// TIA Portal V20 export
TYPE "Afag_Variablen_Steuerung_Dreh"
   STRUCT
      BA_Manuell : Bool;
      Manuell_Geschwindigkeit_in_P : Int := 10;
      Richten_Reset_FRG : Bool;
      drive_enable : Bool;
      start_homing : Bool;
      jog_pos : Bool;
      jog_neg : Bool;
      fault_reset : Bool;
      Tipp_pos : Bool;
      Tipp_neg : Bool;
      Start_pos_man : Bool;
      Verfahrweg_Grad : Real;
      soll_wert_man_Grad : Real;
      Softw_ES_min_Grad : Real;
      Softw_ES_max_Grad : Real;
      Max_Speed_Grad_s : Real;
      Max_Beschleunigung_Grad_s : Real;
      drive_enable_ok : Bool;
      home_valid : Bool;
      pos_ok : Bool;
      velo_zero : Bool;
      fault : Bool;
      Positionsfehler : Bool;
      Fahrauftrag_Aktiv : Bool;
      ist_wert_Grad : Real;
   END_STRUCT;
END_TYPE
